// Mitsubishi GX Works2 project: Practica d   PLC: FX3G

PROGRAM MAIN
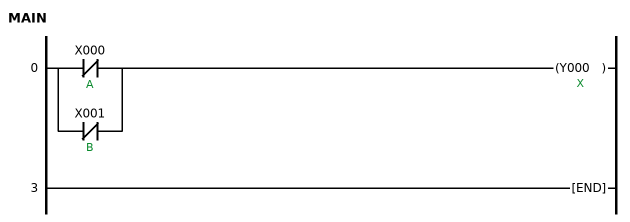
0     LDI     X000  ; A
      ORI     X001  ; B
      OUT     Y000  ; X
3     END
END_PROGRAM
